Staubli VAL3: Lab2B_L3.dtx


